// TIA Portal V20 export
Screen "Pop-up_ATDC"  395x500
  ScreenItem "Robot Name" at 2,2 size 393x48  Type=HmiIOField
  ScreenItem "Background" at -1,49 size 395x450  Type=HmiRectangle
  ScreenItem "Cancel Mode" at 315,4 size 76x42  Type=HmiButton
  ScreenItem "矩形_4" at 29,63 size 324x402  Type=HmiRectangle
  ScreenItem "Text Filed E- Stop_17" at 41,339 size 298x21  Type=HmiTextBox
  ScreenItem "Text Field In Auto On_9" at 41,99 size 298x21  Type=HmiTextBox
  ScreenItem "Text Field Home Position_17" at 41,123 size 298x21  Type=HmiTextBox
  ScreenItem "Text field Robot Status_5" at 31,64 size 324x30  Type=HmiTextBox
  ScreenItem "Text Field Manual_17" at 41,267 size 298x21  Type=HmiTextBox
  ScreenItem "Text Field System Ready_9" at 41,147 size 298x21  Type=HmiTextBox
  ScreenItem "Text Field Motor On_9" at 41,171 size 298x21  Type=HmiTextBox
  ScreenItem "Text Field In Cycle_9" at 41,195 size 298x21  Type=HmiTextBox
  ScreenItem "Text Field Cycle On_17" at 41,219 size 298x21  Type=HmiTextBox
  ScreenItem "Text Field On Path_17" at 41,243 size 298x21  Type=HmiTextBox
  ScreenItem "Text Field Tryout Mode_17" at 41,291 size 298x21  Type=HmiTextBox
  ScreenItem "Text Field Stop_17" at 41,315 size 298x21  Type=HmiTextBox
  ScreenItem "Text Filed Error_9" at 41,363 size 298x21  Type=HmiTextBox
  ScreenItem "Text Filed Process Fault_9" at 41,387 size 298x21  Type=HmiTextBox
  ScreenItem "Text Filed Process Fault_1" at 41,411 size 298x21  Type=HmiTextBox
  ScreenItem "Text Filed Process Fault_2" at 41,434 size 298x21  Type=HmiTextBox
